(* IEC 61131-3 sources: POMIRTS_lab3/AS/Library_2/AsMbTCPS, 3 files *)

(* ---- AsMbTCPS.typ ---- *)
TYPE

END_TYPE

(* ---- AsMbTCPS.fun ---- *)
{REDUND_CONTEXT} {REDUND_UNREPLICABLE} FUNCTION_BLOCK mbSlBoolPut							(*writes bit-oriented slave data; synchronous execution*)
	VAR_INPUT
		enable			: BOOL;						(*enables execution*)
		startAddress	: UINT;						(*starting address*)
		nrOfItems		: USINT;						(*number of items to write*)
	END_VAR

	VAR_IN_OUT
		station			: STRING[1]; 				(*station path e.g."IF2.MODBUSSLAVE_1"*)
		data			: ARRAY[0..127] OF BOOL;	(*array of data, only the first "nrOfItems" will be used*)
	END_VAR

	VAR
	END_VAR

	VAR_OUTPUT
		status			: UINT;						(*execution status: ERR_OK, ERR_FUB_ENABLE_FALSE, 0xXXXX = see help*)
	END_VAR
END_FUNCTION_BLOCK

{REDUND_CONTEXT} {REDUND_UNREPLICABLE} FUNCTION_BLOCK mbSlBoolGet							(*reads bit-oriented slave data; synchronous execution*)
	VAR_INPUT
		enable			: BOOL;						(*enables execution*)
		startAddress	: UINT;						(*starting address*)
		nrOfItems		: USINT;						(*number of items to read*)
	END_VAR

	VAR_IN_OUT
		station			: STRING[1]; 				(*station path e.g."IF2.MODBUSSLAVE_1"*)
		data			: ARRAY[0..127] OF BOOL;	(*array which will be filled with the requested data*)
	END_VAR

	VAR
	END_VAR

	VAR_OUTPUT
		status			: UINT;						(*execution status: ERR_OK, ERR_FUB_ENABLE_FALSE, 0xXXXX = see help*)
	END_VAR
END_FUNCTION_BLOCK

{REDUND_CONTEXT} {REDUND_UNREPLICABLE} FUNCTION_BLOCK mbSlWordPut							(*writes word-oriented slave data; synchronous execution*)
	VAR_INPUT
		enable			: BOOL;						(*enables execution*)
		startAddress	: UINT;						(*starting address*)
		nrOfItems		: USINT;						(*number of items to write*)
	END_VAR

	VAR_IN_OUT
		station			: STRING[1]; 				(*station path e.g."IF2.MODBUSSLAVE_1"*)
		data			: ARRAY[0..127] OF UINT;	(*array of data*)
	END_VAR

	VAR
	END_VAR

	VAR_OUTPUT
		status			: UINT;						(*execution status: ERR_OK, ERR_FUB_ENABLE_FALSE, 0xXXXX = see help*)
	END_VAR
END_FUNCTION_BLOCK

{REDUND_CONTEXT} {REDUND_UNREPLICABLE} FUNCTION_BLOCK mbSlWordGet							(*reads word-oriented slave data; synchronous execution*)
	VAR_INPUT
		enable			: BOOL;						(*enables execution*)
		startAddress	: UINT;						(*starting address*)
		nrOfItems		: USINT;						(*number of items to read*)
	END_VAR

	VAR_IN_OUT
		station			: STRING[1]; 				(*station path e.g."IF2.MODBUSSLAVE_1"*)
		data			: ARRAY[0..127] OF UINT;	(*array which will be filled with the requested data*)
	END_VAR

	VAR
	END_VAR

	VAR_OUTPUT
		status			: UINT;						(*execution status: ERR_OK, ERR_FUB_ENABLE_FALSE, 0xXXXX = see help*)
	END_VAR
END_FUNCTION_BLOCK

(* ---- AsMbTCPS.var ---- *)
VAR CONSTANT
	mbSlOFFSET_DISCRETE_INPUT			: UINT := 0;			(*startaddress of discrete input addressspace => 0x0000*)
	mbSlOFFSET_COIL						: UINT := 16384;		(*startaddress of coil addressspace => 0x4000*)
	mbSlOFFSET_INPUT_REGISTER			: UINT := 8192;			(*startaddress of coil addressspace => 0x2000*)
	mbSlOFFSET_HOLDING_REGISTER			: UINT := 24576;		(*startaddress of coil addressspace => 0x6000*)
	mbSlERR_INVALID_CONFIG				: UINT := 37450;		(*slave has to be configured with fixed buffersize*)
	mbSlERR_INVALID_STATION				: UINT := 37451;		(*station does not exist*)
	mbSlERR_INVALID_ADDRESS				: UINT := 37452;		(*startaddress or number of coils/registers incorrect*)
	mbSlERR_NULLPOINTER					: UINT := 37453;		(*nullpointer*)
	mbSlERR_INVALID_NUMBER_OF_ITEMS		: UINT := 37454;		(*Number of Items must be between 1 and 128*)
END_VAR
